Fanuc KAREL source: kb00042.KL

-- PROVISIONAL review KL for V770-1; original PC SHA256 e0f9b22b66ae1f36ef262ff5a47d8c9758b0352a0a06c9be0340a00f29667460
-- Incomplete behavior may be omitted. Consult companion uncertainty JSON. Do not deploy.
PROGRAM KB00042
%NOLOCKGROUP
BEGIN
  -- UNRESOLVED_PC offsets 5-14; opcodes 3F,75
  -- UNRESOLVED_PC offsets 19-26; opcodes 9D,23
  -- UNRESOLVED_PC offsets 31-49; opcodes 27,22,2A,22,31
  -- UNRESOLVED_PC offsets 54-58; opcodes 7F
END KB00042
